(* IEC 61131-3 sources: SortJet_MasterSPS_Aufbau.fbsproj/09_Station/Stationen/Faecherwagen [301-305], 6 files *)

(* ---- I_Faecherwagenstation.itf ---- *)
(* METADATA
{
	"v3Meta": {
		"objectGuid": "03e38843-2da5-4b21-8acb-320ccd699887"
	}
}
*)
INTERFACE I_Faecherwagenstation EXTENDS __System.IQueryInterface
END_INTERFACE

(* ---- Basic_Faecherwagenstation_FB_V01_00_00.fb.st ---- *)
(* METADATA
{
	"v3Meta": {
		"objectGuid": "908407cd-758c-45db-8a2d-c326aeb0e347"
	}
}
*)
FUNCTION_BLOCK ABSTRACT Basic_Faecherwagenstation_FB_V01_00_00 EXTENDS Basic_Station_FB_V01_00_00 IMPLEMENTS I_Faecherwagenstation
VAR_INPUT

  // BOOL
  blMerkerEinschleusenQuittiert     : BOOL; // Einschleusen vom Bediener an der Station quittiert
  bpRolltorUnten                    : BOOL; // Rolltor unten (aus der Sicherheitstechnik)
  bpMMIFWBaldVoll                   : BOOL; // Faecherwagen in der Station laut MMI bald voll (Anzeige an der Station), Ruecksetzen beim Verlassen der Beladeposition

  // WORD
  wlRFID_Nummer_Schreiben           : WORD; // Neue Nummer fuer den RFID-Chip des Faecherwagens (vom MMI)

  // USINT
  usilErrorSafety                   : USINT; // Fehlercode der sicheren Feldbox (Schmersal), im Geraetebaum gemappt

END_VAR
VAR_OUTPUT

  // BOOL
  bpDone                            : BOOL;
  bpEinschleusenAbgeschlossen       : BOOL;
  bpAusschleusenAbgeschlossen       : BOOL;
  bpAuftragAktiv                    : BOOL;
  bpFehler                          : BOOL;
  bpErzwingeAusschleusen            : BOOL;
  bpErzwingeEinschleusen            : BOOL;
  bpBoxInHomePosition               : BOOL; // Mechanik der Station in Grundstellung
  bpOutBereitZumAustransport        : BOOL; // OUT STATUS: Bereit zum Austransport [Eintransport auf die Nachfolgerstation]
  bpOutBereitZumEintransport        : BOOL; // OUT STATUS: Bereit zum Eintransport [Austransport auf die Vorgaengerstation]
  bpStatusStationInBeladePosition   : BOOL; // Faecherwagen steht in der Beladeposition (zyklisch)
  bpHinweisEingriffErforderlich     : BOOL; // Bedienereingriff am Faecherwagen erforderlich (Ampel blau blinkend, Aktion Ampelsignal in Job)

  // WORD
  wpFehlerNr                        : Fehlerkonstanten_EN; // FEHLER-AUSWERTUNG: Fehlernummer[Const]

END_VAR
VAR

  // BOOL
  blRolltorAuf                      : BOOL; // Anforderung Rolltor oeffnen
  blRolltorAb                       : BOOL; // Anforderung Rolltor schliessen
  blRolltorAufDone                  : BOOL;
  blRolltorAbDone                   : BOOL;
  blRolltorAbFreigabe               : BOOL := TRUE; // Variante: Rolltor darf schliessen (z.B. nichts im Bereich des Rolltors)
  blRolltorAbBlockiert              : BOOL; // Variante: Schliessen sofort mit Fehler abbrechen (z.B. Abrollsicherung ausgeloest)
  blStationsposUndefiniert          : BOOL; // Station weder in Grundstellung noch in Beladeposition und kein Auftrag aktiv
  blStarteSicherheitskreisReset     : BOOL; // Anforderung Sicherheitsrelais der Station quittieren (MMI, Variante setzt nach Ausfuehrung zurueck)
  blAckRequested                    : BOOL; // Sichere Feldbox fordert Quittierung an, im Geraetebaum gemappt
  blResetSchmersal                  : BOOL; // Quittierimpuls an die sichere Feldbox, im Geraetebaum gemappt

  // WORD
  wlZeitHochfahren                  : WORD;
  wlZeitRunterfahren                : WORD;
  wlRFID_Nummer                     : WORD; // Zuletzt gelesene RFID-Nummer des Faecherwagens

  // TIME
  tlZeitHochfahren                  : TIME;
  tlZeitRunterfahren                : TIME;

  // STEPS
  steplRolltorAuf                   : Steps_TE;
  steplRolltorAb                    : Steps_TE;

  // TIMER
  tonlFreigabe                      : TON;
  tonlUeberwachungRolltor           : TON;
  tonlRolltorOeffnenSchliesen       : TON;
  tonlZeitRunterfahren              : TON; // Zum ermitteln wie lange das Rolltor runterfaehrt
  tonlZeitHochfahren                : TON; // Zum ermitteln wie lange das Rolltor hochfaehrt
  tplResetSchmersal                 : TP;

  // TRIGGER
  rtlSafetyError                    : R_TRIG;

  // ENUM
  eLetzterStatus                    : eLetzter_FW_Status; // Zuletzt erreichter Schritt fuer Systemcheck und MMI
  elLetzterStatusGesendet           : eLetzter_FW_Status; // Zuletzt ans MMI gemeldeter Status (STATION_UPDATE)

  // HARDWARE: ROLLTOR
  in_bRolltorGeoeffnet                     : BOOL; // TRUE = Rolltor oben, im Geraetebaum gemappt
  out_bRolltorAb                    AT %Q* : BOOL;
  out_bRolltorAuf                   AT %Q* : BOOL;

  // HARDWARE: SICHERHEITSKREIS DER STATION (im Geraetebaum gemappt)
  in_bResetSicherheitskreis         : BOOL; // Taster Sicherheitskreis quittieren an der Station
  out_bSicherheitskreisAusgeloest   : BOOL; // Leuchte Sicherheitskreis ausgeloest (Variante darf ueberschreiben)

END_VAR
VAR CONSTANT

  // TIME
  cZEIT_UEBERWACHUNG_ROLLTOR        : TIME := T#60S;

END_VAR
//-------------------------------------------------------------------------------------------------
// MASTER AUFRUFEN
//-------------------------------------------------------------------------------------------------
IF NOT __ISVALIDREF(BasisStationsParameter.stMKs) THEN
  dwpHandfunktionenReturn := DWORD#0;
  RETURN;
END_IF

SUPER^(BasisStationsParameter := BasisStationsParameter);

//-------------------------------------------------------------------------------------------------
// DEAKTIVIEREN
//-------------------------------------------------------------------------------------------------
// Werte wieder passend abloeschen, wenn der Baustein wieder aktiviert wird
IF ( ftlBausteinDeaktivierung.Q ) THEN
  bpDone                      := FALSE;
  bpEinschleusenAbgeschlossen := FALSE;
  bpAusschleusenAbgeschlossen := FALSE;
END_IF

(* Hinweis:
   - Deaktivierte Station: nichts melden, nichts bewegen
   - Die Variante prueft die Deaktivierung nach dem Aufruf selbst und setzt ihre Anforderungen zurueck
*)
IF ( BasisStationsParameter.stMKs.bDeaktivieren ) THEN

  bpDone                          := TRUE;
  bpEinschleusenAbgeschlossen     := TRUE;
  bpAusschleusenAbgeschlossen     := TRUE;
  bpStatusStationInBeladePosition := FALSE;
  bpAuftragAktiv                  := FALSE;
  bpFehler                        := FALSE;
  blStationsposUndefiniert        := FALSE;

  blRolltorAuf                    := FALSE;
  blRolltorAb                     := FALSE;
  out_bRolltorAuf                 := FALSE;
  out_bRolltorAb                  := FALSE;

  A_Visu();
  RETURN;

END_IF

//-------------------------------------------------------------------------------------------------
// TIMER
//-------------------------------------------------------------------------------------------------
tonlFreigabe( IN := BasisStationsParameter.stFreigabe.bAlles, PT := T#1S );

bpFehler := BasisStationsParameter.bFehler;

//-------------------------------------------------------------------------------------------------
// SICHERE FELDBOX / SICHERHEITSKREIS
//-------------------------------------------------------------------------------------------------
rtlSafetyError( CLK := usilErrorSafety <> 0 );
IF rtlSafetyError.Q THEN

  SpsError( eFehler_Safety_Schmersal,
            usilErrorSafety,
            BasisStationsParameter.stMKs.stStationsNummern.NummerIntern,
            AutomatikkreisBestimmen(BasisStationsParameter.stMKs.stStationsNummern.NummerSPS),
            BasisStationsParameter.awFehlerInformationen );

END_IF

tplResetSchmersal( IN := blAckRequested XOR ( NotHalt.in_bTasterNothaltQuittieren OR in_bResetSicherheitskreis ),
                   PT := T#500MS,
                   Q  => blResetSchmersal );

// Meldung "Faecherwagen bald voll" gilt nur fuer den Faecherwagen in der Beladeposition
IF NOT bpStatusStationInBeladePosition THEN
  bpMMIFWBaldVoll := FALSE;
END_IF

//-------------------------------------------------------------------------------------------------
// STATUS AN MMI MELDEN
//-------------------------------------------------------------------------------------------------
// Hinweis:
//   - Der fuer den Systemcheck gemerkte Status (eLetzterStatus) wird bei jeder Aenderung und bei
//     neuer MMI-Verbindung gemeldet; das MMI zeigt die Geraete der Station passend dazu an
IF ( eLetzterStatus <> elLetzterStatusGesendet ) OR Job.rtlMmiOk.Q THEN
  stStationUpdate.wStationsNummer       := BasisStationsParameter.stMKs.stStationsNummern.NummerSPS;
  stStationUpdate.eUpdateTyp            := StationUpdateTyp_EN.FW_STATUS;
  stStationUpdate.wAnzahlWerte          := 1;
  stStationUpdate.astWerte[1].eDatenTyp := UpdateDatenTyp_EN.TYP_WORD;
  stStationUpdate.astWerte[1].wWert     := TO_WORD( eLetzterStatus );
  MsgToMmi( auftragsnr_w := SB0_SPS_STATION_UPDATE );

  elLetzterStatusGesendet := eLetzterStatus;
END_IF
END_FUNCTION_BLOCK

(* ---- Faecherwagenstation_Einfach_FB_V01_00_00.fb.st ---- *)
(* METADATA
{
	"v3Meta": {
		"objectGuid": "602268ae-05d1-404e-8d8e-505fe92152ba"
	}
}
*)
FUNCTION_BLOCK Faecherwagenstation_Einfach_FB_V01_00_00 EXTENDS Basic_Faecherwagenstation_FB_V01_00_00
VAR_INPUT

  // BOOL
  bpFaecherwagenVorhanden          : BOOL; // Faecherwagen vorhanden, Sicherheitssensor ueber die SLC (Interface_SLC)
  in_bDruckluftOK                  : BOOL;

END_VAR
VAR

  // BOOL
  blArretierungSchliessen          : BOOL; // Anforderung Arretierung ausfahren (Faecherwagen festhalten)
  blArretierungOeffnen             : BOOL; // Anforderung Arretierung einfahren (Faecherwagen freigeben)
  blArretierungSchliessenDone      : BOOL;
  blArretierungOeffnenDone         : BOOL;
  blArretierungGeschlossen         : BOOL; // Arretierung ausgefahren (Endlage)
  blArretierungOffen               : BOOL; // Arretierung eingefahren (Endlage)
  blHandFreigabe                   : BOOL; // Handfunktionen nur im Handbetrieb zulassen
  blTasterLeuchteAnforderung       : BOOL;

  // WORD
  wlIoccMeldungsNummer             : WORD;

  // STEPS
  steplEinschleusen                : Steps_TE;
  steplAusschleusen                : Steps_TE;

  // TIMER
  tonlFWInBox                      : TON; // Faecherwagen steht stabil in der Station
  tonlErzwungenesAuschleusen       : TON;

  // TRIGGER
  rtlLogIn                         : R_TRIG;
  rtlQuittierungEinschleusen       : R_TRIG;
  rtlBetriebsartHand               : R_TRIG;
  ftlBetriebsartAutomatik          : F_TRIG;
  rtlArretierungFehler             : R_TRIG;

  // BAUSTEINE
  Arretierung                      : Arretierung_FB_V01_00_00; // Arretierung (Zentrierung/Klemmung) des ganzen Faecherwagens

  // HARDWARE EINGAENGE (Konfiguration_FW_Einfach)
  in_bAbrollsicherungOK            AT %I* : BOOL; // Abrollsicherung am Rolltor in Ordnung (Oeffner: TRUE = frei)

  // HARDWARE EINGAENGE (IO-Link, im Geraetebaum gemappt)
  in_bArretierungAusgefahren       : BOOL; // Faecherwagen arretiert
  in_bArretierungEingefahren       : BOOL; // Faecherwagen freigegeben
  in_bStartSchleusen               : BOOL; // Taster Ein-/Ausschleusen an der Station

  // HARDWARE AUSGAENGE (IO-Link, im Geraetebaum gemappt)
  out_bArretierungAusfahren        : BOOL;
  out_bArretierungEinfahren        : BOOL;
  out_bFreigabeSchleusen           : BOOL; // Leuchte im Taster Ein-/Ausschleusen

END_VAR
VAR CONSTANT

  // TIME
  ZEIT_ZWANGSAUSSCHLEUSEN          : TIME := T#3S;
  ZEIT_FW_IN_BOX                   : TIME := T#2S;

END_VAR

//-------------------------------------------------------------------------------------------------
// MASTER AUFRUFEN
//-------------------------------------------------------------------------------------------------
IF NOT __ISVALIDREF(BasisStationsParameter.stMKs) THEN
  dwpHandfunktionenReturn := DWORD#0;
  RETURN;
END_IF

SUPER^(BasisStationsParameter := BasisStationsParameter);

//-------------------------------------------------------------------------------------------------
// DEAKTIVIEREN
//-------------------------------------------------------------------------------------------------
IF ( BasisStationsParameter.stMKs.bDeaktivieren ) THEN

  blArretierungSchliessen   := FALSE;
  blArretierungOeffnen      := FALSE;
  out_bArretierungAusfahren := FALSE;
  out_bArretierungEinfahren := FALSE;
  out_bFreigabeSchleusen    := FALSE;

  HandfunktionenStatus();
  RETURN;

END_IF

//-------------------------------------------------------------------------------------------------
// AKTIONEN
//-------------------------------------------------------------------------------------------------
A_Eingaenge();
Ausschleusen();
Einschleusen();
Rolltor();

Systemcheck();

Reset();
Handfunktionen();

A_Aufrufe();
Ausgaenge();

A_Visu();
A_VisuVariante();

//-------------------------------------------------------------------------------------------------
// TASTER
//-------------------------------------------------------------------------------------------------
IF BasisStationsParameter.bEintransport[cWAND_1] THEN

  IF steplEinschleusen = STEP_105_E THEN
    blTasterLeuchteAnforderung := gbFlashbit05sec; // Einschleusen wartet auf die Quittierung
  ELSE
    blTasterLeuchteAnforderung := gbFlashbit1sec;
  END_IF

ELSIF BasisStationsParameter.bAustransport[cWAND_1] THEN
  blTasterLeuchteAnforderung := gbFlashbit1sec;

ELSIF blStationsposUndefiniert THEN
  blTasterLeuchteAnforderung := gbFlashbit02sec; // Undefinierter Zustand - sehr schnell blinken

ELSIF bpStatusStationInBeladePosition THEN
  blTasterLeuchteAnforderung := bpMMIFWBaldVoll; // Faecherwagen in Beladeposition: Dauerlicht, wenn er laut MMI bald voll ist

ELSIF bpBoxInHomePosition THEN
  blTasterLeuchteAnforderung := TRUE; // Station bereit zum Einschleusen

ELSE
  blTasterLeuchteAnforderung := gbFlashbit02sec;
END_IF

out_bFreigabeSchleusen := blTasterLeuchteAnforderung;

//-------------------------------------------------------------------------------------------------
// GESONDERTE LOGIK
//-------------------------------------------------------------------------------------------------

// Ausschleusen erzwingen: Taster lange druecken
tonlErzwungenesAuschleusen( IN := in_bStartSchleusen, PT := ZEIT_ZWANGSAUSSCHLEUSEN );
bpErzwingeAusschleusen := tonlErzwungenesAuschleusen.Q;

// Faecherwagen anmelden: Taster bei Faecherwagen in der Station und Station in Grundstellung
rtlLogIn( CLK :=     in_bStartSchleusen
                 AND bpBoxInHomePosition
                 AND tonlFWInBox.Q
                 AND NOT bpStatusStationInBeladePosition
                 AND NOT bpAuftragAktiv );

IF ( rtlLogIn.Q ) THEN
  wSps2FaecherwagenStationNr              := BasisStationsParameter.stMKs.stStationsNummern.NummerSPS;
  tMmi2SpsInfo.wSps2FaecherwagenStationNr := BasisStationsParameter.stMKs.stStationsNummern.NummerSPS;
  MsgToMmi( auftragsnr_w := SB0_SPS_RACKLOGIN );

  M_SB0_MMI_RELEASERACKLOGIN    := TRUE;
  blMerkerEinschleusenQuittiert := TRUE;
END_IF
END_FUNCTION_BLOCK

(* ---- Faecherwagenstation_Hydraulik_FB_V01_00_00.fb.st ---- *)
(* METADATA
{
	"v3Meta": {
		"objectGuid": "e6879d41-371d-40de-a0ee-fe2898e6d6d8"
	}
}
*)
FUNCTION_BLOCK Faecherwagenstation_Hydraulik_FB_V01_00_00 EXTENDS Basic_Faecherwagenstation_FB_V01_00_00
VAR_OUTPUT

  // BOOL
  bpAnforderungHydraulikEin        : BOOL; // Hydraulikaggregat einschalten (eine hydraulische Bewegung ist angefordert)
  bpUmlaufVentilPause              : BOOL; // Umlaufventil zwischen zwei direkt folgenden Bewegungen kurz zuruecknehmen

END_VAR
VAR

  // BOOL: Anforderungen
  blHubrahmenHeben                 : BOOL;
  blHubrahmenSenken                : BOOL;
  blFaecherwagenVor                : BOOL;
  blFaecherwagenZurueck            : BOOL;
  blZentrierungOeffnen             : BOOL;
  blZentrierungSchliessen          : BOOL;
  blAnschlagAuf                    : BOOL;
  blAnschlagAb                     : BOOL;
  blAnschlagVor                    : BOOL; // Option AGV: Anschlag nach vorne
  blAnschlagZurueck                : BOOL; // Option AGV: Anschlag nach hinten

  // BOOL: Bewegungen abgeschlossen
  blHubrahmenHebenDone             : BOOL;
  blHubrahmenSenkenDone            : BOOL;
  blFaecherwagenVorDone            : BOOL;
  blFaecherwagenZurueckDone        : BOOL;
  blZentrierungOeffnenDone         : BOOL;
  blZentrierungSchliessenDone      : BOOL;
  blAnschlagAufDone                : BOOL;
  blAnschlagAbDone                 : BOOL;
  blAnschlagVorDone                : BOOL;
  blAnschlagZurueckDone            : BOOL;

  // BOOL: Verschiedenes
  blFaecherwagenErkannt            : BOOL; // Beide Muting-Sensoren belegt
  blAnschlagUntenOderOhne          : BOOL; // Anschlag unten oder kein Anschlag laut MK
  blLadepositionOhneOben           : BOOL; // Beladeposition bis auf den abgesackten Hubrahmen
  blPositionskorrekturAktiv        : BOOL; // Hubrahmen wird nachgehoben
  blAnforderungHydraulik           : BOOL;
  blHandFreigabe                   : BOOL; // Handfunktionen nur im Handbetrieb zulassen
  blTasterLeuchteAnforderung       : BOOL;
  blHydraulikLaeuft                : BOOL; // Rueckmeldung der zugeordneten Hydraulikstation
  blStationBeladen                 : BOOL; // Faecherwagen eingeschleust (Status fuer AGV-Betrieb)
  blStartUp                        : BOOL := TRUE; // Sicherheitsrelais nach dem Programmstart einmal quittieren

  // BOOL: Begrenzung gleichzeitiger Auftraege je Hydraulikstation
  blHydraulikAuftragAnfrage        : BOOL; // Kette wartet auf die Freigabe eines neuen Auftrags (je Zyklus neu gesetzt)
  blHydraulikAuftragFreigabe       : BOOL; // Rueckmeldung der Hydraulikstation (M_AuftragFreigabe, letzter Zyklus)
  blHydraulikAuftragAktiv          : BOOL; // Ein-/Ausschleusen mit hydraulischen Bewegungen laeuft, belegt die Hydraulikstation
  blAuftragWartetAufHydraulik      : BOOL; // Auftrag erteilt, Hydraulikstation laesst noch keinen weiteren Auftrag zu

  // BOOL: Muting
  blMutingAusschalten              : BOOL; // Option AGV: Muting dauerhaft zuruecksetzen (kein Faecherwagen eingeschleust)
  blMutingResetAnforderung         : BOOL; // Anforderung Muting-Sensoren zuruecksetzen pruefen
  blMutingResetImpuls              : BOOL; // Reset-Impuls fuer die Muting-Sensoren ausgeben
  blMutingSensorReset              : BOOL; // Reset-Impuls aktiv

  // BYTE
  bylRFID_Nummer                   : BYTE;

  // WORD
  wlIoccMeldungsNummer             : WORD;
  wlStationStatusWord              : WORD; // Option AGV: zuletzt ans MMI gemeldeter Status der Station

  // REFERENZ
  refHydraulikstation              : REFERENCE TO Hydraulik_FB_V01_00_00; // laut MK stStationsAufbau.wHydraulikstation

  // STEPS
  steplEinschleusen                : Steps_TE;
  steplAusschleusen                : Steps_TE;
  steplHubrahmenHeben              : Steps_TE;
  steplHubrahmenSenken             : Steps_TE;
  steplFaecherwagenVor             : Steps_TE;
  steplFaecherwagenZurueck         : Steps_TE;
  steplZentrierungOeffnen          : Steps_TE;
  steplZentrierungSchliessen       : Steps_TE;
  steplSicherheitskreisReset       : Steps_TE;

  // TIMER
  tonlHubrahmenUeberfahren         : TON; // Sensor ueberfahren, Endlage sicher erreicht
  tonlVerfahrenUeberfahren         : TON;
  tonlZentrierungUeberfahren       : TON;
  tonlTimeoutHubrahmen             : TON;
  tonlTimeoutVerfahren             : TON;
  tonlTimeoutZentrierung           : TON;
  tonlTimeoutHydraulik             : TON; // Warten auf das Hydraulikaggregat
  tonlTimeoutReadRFID              : TON;
  tonlFWInBox                      : TON;
  tonlErzwungenesAuschleusen       : TON;
  tonlMutingSensorFehler           : TON;
  tonlPositionskorrektur           : TON;
  tonlUmlaufventilPause            : TON; // Dauer der Pause des Umlaufventils
  tonlMutingSensorenBelegt         : TON; // Beide Muting-Sensoren stabil belegt
  tonlTimeoutAGV                   : TON; // Option AGV: Warten auf den Faecherwagen
  tonlRFIDGelesen                  : TON; // Option AGV: RFID-Chip stabil gelesen
  tonlStartUp                      : TON;
  tonlResetImpuls                  : TON; // Impulsdauer Reset Sicherheitsrelais
  tonlResetWarten                  : TON; // Wartezeiten der Kette Sicherheitskreis-Reset
  toflAnforderungHydraulikEin      : TOF;
  toflMutingSensorReset            : TOF; // Impulsdauer Reset Muting-Sensoren

  // TRIGGER
  rtlLogIn                         : R_TRIG;
  rtlQuittierungEinschleusen       : R_TRIG;
  rtlBetriebsartHand               : R_TRIG;
  ftlBetriebsartAutomatik          : F_TRIG;
  rtlPositionskorrektur            : R_TRIG;
  rtlAnschlagFehler                : R_TRIG;
  rtlAnschlagHorizontalFehler      : R_TRIG;
  rtlMutingSensorReset             : R_TRIG;
  ftlRFIDNichtMehrGelesen          : F_TRIG;

  // BAUSTEINE
  Anschlag                         : ZylinderPneumatik_FB_V01_00_00; // Option stStationsAufbau.bAnschlag, ausgefahren = oben
  AnschlagHorizontal               : ZylinderPneumatik_FB_V01_00_00; // Option bAnschlag und bAGV, ausgefahren = vorne

  // HARDWARE EINGAENGE
  in_bHubrahmenOben                AT %I* : BOOL;
  in_bHubrahmenUnten               AT %I* : BOOL;
  in_bFaecherwagenVorne            AT %I* : BOOL;
  in_bFaecherwagenHinten           AT %I* : BOOL;
  in_bZentrierungOffen             AT %I* : BOOL;
  in_bZentrierungGeschlossen       AT %I* : BOOL;
  in_bAnschlagOben                 AT %I* : BOOL;
  in_bAnschlagUnten                AT %I* : BOOL;
  in_bAnschlagVorne                AT %I* : BOOL; // Option AGV
  in_bAnschlagHinten               AT %I* : BOOL; // Option AGV
  in_bFWInAusrichtPosition         AT %I* : BOOL; // Faecherwagen steht vor der Station in Ausrichtposition
  in_bMutingSensorLinks            AT %I* : BOOL;
  in_bMutingSensorRechts           AT %I* : BOOL;
  in_bStartSchleusen               AT %I* : BOOL; // Taster Ein-/Ausschleusen an der Station
  in_bSicherheitsrelaisOK          AT %I* : BOOL;
  in_bAbrollsicherungOK            AT %I* : BOOL; // Abrollsicherung des Rolltors nicht ausgeloest
  in_bRFID_DataValid               AT %I* : BOOL;
  in_bRFID_NR1                     AT %I* : BOOL;
  in_bRFID_NR2                     AT %I* : BOOL;
  in_bRFID_NR3                     AT %I* : BOOL;
  in_bRFID_NR4                     AT %I* : BOOL;
  in_bRFID_NR5                     AT %I* : BOOL;
  in_bRFID_NR6                     AT %I* : BOOL;
  in_bRFID_NR7                     AT %I* : BOOL;
  in_bRFID_NR8                     AT %I* : BOOL;

  // HARDWARE AUSGAENGE
  out_bHubrahmenHeben              AT %Q* : BOOL;
  out_bHubrahmenSenken             AT %Q* : BOOL;
  out_bFaecherwagenVor             AT %Q* : BOOL;
  out_bFaecherwagenZurueck         AT %Q* : BOOL;
  out_bZentrierungOeffnen          AT %Q* : BOOL;
  out_bZentrierungSchliessen       AT %Q* : BOOL;
  out_bAnschlagAuf                 AT %Q* : BOOL;
  out_bAnschlagAb                  AT %Q* : BOOL;
  out_bAnschlagVor                 AT %Q* : BOOL; // Option AGV
  out_bAnschlagZurueck             AT %Q* : BOOL; // Option AGV
  out_bFreigabeSchleusen           AT %Q* : BOOL; // Leuchte im Taster Ein-/Ausschleusen
  out_bMutingSensorReset           AT %Q* : BOOL; // Muting-Sensoren zuruecksetzen
  out_bResetSicherheitsrelais      AT %Q* : BOOL; // Sicherheitsrelais der Station quittieren

END_VAR
VAR CONSTANT

  // TIME
  ZEIT_TIMEOUT_SENSOR              : TIME := T#30S;
  ZEIT_TIMEOUT_HYDRAULIK           : TIME := T#30S;
  ZEIT_SENSOR_UEBERFAHREN          : TIME := T#3S;
  ZEIT_POSITIONSKORREKTUR          : TIME := T#5S;
  ZEIT_TIMEOUT_RFID                : TIME := T#5S;
  ZEIT_ZWANGSAUSSCHLEUSEN          : TIME := T#3S;
  ZEIT_FW_IN_BOX                   : TIME := T#1S;
  ZEIT_UMLAUFVENTIL_PAUSE          : TIME := T#1S;
  ZEIT_MUTING_SENSOR_RESET         : TIME := T#500MS;
  ZEIT_STARTUP_SICHERHEITSRELAIS   : TIME := T#5S;

END_VAR
//-------------------------------------------------------------------------------------------------
// MASTER AUFRUFEN
//-------------------------------------------------------------------------------------------------
IF NOT __ISVALIDREF(BasisStationsParameter.stMKs) THEN
  dwpHandfunktionenReturn := DWORD#0;
  RETURN;
END_IF

SUPER^(BasisStationsParameter := BasisStationsParameter);

//-------------------------------------------------------------------------------------------------
// DEAKTIVIEREN
//-------------------------------------------------------------------------------------------------
IF ( BasisStationsParameter.stMKs.bDeaktivieren ) THEN

  blHubrahmenHeben           := FALSE;
  blHubrahmenSenken          := FALSE;
  blFaecherwagenVor          := FALSE;
  blFaecherwagenZurueck      := FALSE;
  blZentrierungOeffnen       := FALSE;
  blZentrierungSchliessen    := FALSE;
  blAnschlagAuf              := FALSE;
  blAnschlagAb               := FALSE;
  blAnschlagVor              := FALSE;
  blAnschlagZurueck          := FALSE;
  blPositionskorrekturAktiv  := FALSE;
  blMutingResetImpuls        := FALSE;
  steplSicherheitskreisReset := STEP_0_E;

  out_bHubrahmenHeben        := FALSE;
  out_bHubrahmenSenken       := FALSE;
  out_bFaecherwagenVor       := FALSE;
  out_bFaecherwagenZurueck   := FALSE;
  out_bZentrierungOeffnen    := FALSE;
  out_bZentrierungSchliessen := FALSE;
  out_bAnschlagAuf           := FALSE;
  out_bAnschlagAb             := FALSE;
  out_bAnschlagVor            := FALSE;
  out_bAnschlagZurueck        := FALSE;
  out_bFreigabeSchleusen      := FALSE;
  out_bMutingSensorReset      := FALSE;
  out_bResetSicherheitsrelais := FALSE;
  bpAnforderungHydraulikEin   := FALSE;
  bpUmlaufVentilPause         := FALSE;

  HandfunktionenStatus();
  RETURN;

END_IF

//-------------------------------------------------------------------------------------------------
// AKTIONEN
//-------------------------------------------------------------------------------------------------
A_Eingaenge();
Ausschleusen();
Einschleusen();
Positionskorrektur();

Hubrahmen();
Verfahren();
Zentrierung();
Rolltor();

Systemcheck();
Status_Meldung();

Reset();
Handfunktionen();

MutingSensorReset();
Sicherheitskreis_Reset();

A_Aufrufe();
Ausgaenge();

A_Visu();
A_VisuVariante();

//-------------------------------------------------------------------------------------------------
// TASTER
//-------------------------------------------------------------------------------------------------
IF blAuftragWartetAufHydraulik THEN
  blTasterLeuchteAnforderung := gbFlashbit02sec; // Auftrag erteilt, wartet auf die Hydraulikstation - sehr schnell blinken

ELSIF BasisStationsParameter.bEintransport[cWAND_1] THEN

  IF steplEinschleusen = STEP_100_E THEN
    blTasterLeuchteAnforderung := gbFlashbit05sec; // Einschleusen wartet auf die Quittierung
  ELSE
    blTasterLeuchteAnforderung := gbFlashbit1sec;
  END_IF

ELSIF BasisStationsParameter.bAustransport[cWAND_1] THEN
  blTasterLeuchteAnforderung := gbFlashbit1sec;

ELSIF blStationsposUndefiniert THEN
  blTasterLeuchteAnforderung := gbFlashbit02sec; // Undefinierter Zustand - sehr schnell blinken

ELSIF bpStatusStationInBeladePosition THEN
  blTasterLeuchteAnforderung := bpMMIFWBaldVoll; // Faecherwagen in Beladeposition: Dauerlicht, wenn er laut MMI bald voll ist

ELSIF bpBoxInHomePosition AND in_bFWInAusrichtPosition THEN
  blTasterLeuchteAnforderung := TRUE; // Faecherwagen steht bereit zum Einschleusen

ELSE
  blTasterLeuchteAnforderung := FALSE;
END_IF

out_bFreigabeSchleusen := blTasterLeuchteAnforderung;

//-------------------------------------------------------------------------------------------------
// GESONDERTE LOGIK
//-------------------------------------------------------------------------------------------------

// Ausschleusen erzwingen: Taster lange druecken
tonlErzwungenesAuschleusen( IN := in_bStartSchleusen, PT := ZEIT_ZWANGSAUSSCHLEUSEN );
bpErzwingeAusschleusen := tonlErzwungenesAuschleusen.Q;

// Faecherwagen anmelden: Taster bei Faecherwagen in Ausrichtposition und Station in Grundstellung
rtlLogIn( CLK :=     in_bStartSchleusen
                 AND bpBoxInHomePosition
                 AND tonlFWInBox.Q
                 AND NOT bpStatusStationInBeladePosition
                 AND NOT bpAuftragAktiv );

IF ( rtlLogIn.Q ) THEN
  wSps2FaecherwagenStationNr              := BasisStationsParameter.stMKs.stStationsNummern.NummerSPS;
  tMmi2SpsInfo.wSps2FaecherwagenStationNr := BasisStationsParameter.stMKs.stStationsNummern.NummerSPS;
  MsgToMmi( auftragsnr_w := SB0_SPS_RACKLOGIN );

  M_SB0_MMI_RELEASERACKLOGIN    := TRUE;
  blMerkerEinschleusenQuittiert := TRUE;
END_IF

// Hydraulikaggregat einschalten, solange eine hydraulische Bewegung angefordert und nicht fertig ist
blAnforderungHydraulik :=     BasisStationsParameter.stFreigabe.bAlles
                          AND (    ( blHubrahmenHeben        AND NOT blHubrahmenHebenDone )
                                OR ( blHubrahmenSenken       AND NOT blHubrahmenSenkenDone )
                                OR ( blFaecherwagenVor       AND NOT blFaecherwagenVorDone )
                                OR ( blFaecherwagenZurueck   AND NOT blFaecherwagenZurueckDone )
                                OR ( blZentrierungOeffnen    AND NOT blZentrierungOeffnenDone )
                                OR ( blZentrierungSchliessen AND NOT blZentrierungSchliessenDone ) );

toflAnforderungHydraulikEin( IN := blAnforderungHydraulik, PT := T#2S );
bpAnforderungHydraulikEin := toflAnforderungHydraulikEin.Q;

// Anforderung an die zugeordnete Hydraulikstation melden (Aufruf der Hydraulikstation nach den Faecherwagenstationen)
IF __ISVALIDREF(refHydraulikstation) THEN
  refHydraulikstation.M_Anfordern( bpHydraulikEin      := bpAnforderungHydraulikEin,
                                   bpUmlaufventilPause := bpUmlaufVentilPause );
  blHydraulikLaeuft := refHydraulikstation.bpHydraulikLaeuft;
ELSE
  // Keine Hydraulikstation zugeordnet: hydraulische Bewegungen laufen in die Zeitueberwachung
  blHydraulikLaeuft := FALSE;
END_IF

// Begrenzung gleichzeitiger Auftraege je Hydraulikstation (MK wMaximaleAnzahlAktiverAuftraege):
// Auftrag belegt die Hydraulikstation, bis Ein-/Austransport beendet oder abgebrochen ist
IF     NOT BasisStationsParameter.bEintransport[cWAND_1]
   AND NOT BasisStationsParameter.bAustransport[cWAND_1]
THEN
  blHydraulikAuftragAktiv := FALSE;
END_IF

IF __ISVALIDREF(refHydraulikstation) THEN
  blHydraulikAuftragFreigabe := refHydraulikstation.M_AuftragFreigabe( bpAuftragAktiv   := blHydraulikAuftragAktiv OR blPositionskorrekturAktiv,
                                                                       bpAuftragStarten := blHydraulikAuftragAnfrage );
ELSE
  // Keine Hydraulikstation zugeordnet: keine Begrenzung
  blHydraulikAuftragFreigabe := TRUE;
END_IF

blAuftragWartetAufHydraulik := blHydraulikAuftragAnfrage AND NOT blHydraulikAuftragFreigabe;
blHydraulikAuftragAnfrage   := FALSE;

// Sicherheitsrelais der Station nach dem Programmstart einmal quittieren, sobald Not-Halt in Ordnung ist
tonlStartUp( IN := blStartUp AND NotHalt.bpNotHaltOK, PT := ZEIT_STARTUP_SICHERHEITSRELAIS );

IF ( tonlStartUp.Q ) THEN
  blStartUp                     := FALSE;
  blStarteSicherheitskreisReset := TRUE;
END_IF
END_FUNCTION_BLOCK

(* ---- Faecherwagenstation_Lineareinheit_FB_V01_00_00.fb.st ---- *)
(* METADATA
{
	"v3Meta": {
		"objectGuid": "3779c208-854f-4c13-8b26-aa1147fe8cdb"
	}
}
*)
FUNCTION_BLOCK Faecherwagenstation_Lineareinheit_FB_V01_00_00 EXTENDS Basic_Faecherwagenstation_FB_V01_00_00
VAR_INPUT

  // BOOL
  bpLichtschranke_OK                      : BOOL;// Eingang aus der Sicherheitsteechnik das die Lichtschrnake quittiert ist
  bpUntergestellErkannt                   : BOOL;//safety eingang der Anzeigt, ob ein Unterwagen erkannt wurde
  in_bDruckluftOK                         : BOOL;
  bpLichtschrankeWartetAufQuittierungAmOP : BOOL;

END_VAR
VAR

  //Startet eine Bewegung
  blLineareinheitVor               : BOOL;
  blLineareinheitZurueck           : BOOL;
  blLineareinheitShuttle           : BOOL;
  blEntriegelungOeffnen            : BOOL;
  blEntriegelungSchliessen         : BOOL;
  blGegenhalterOeffnen             : BOOL;
  blGegenhalterSchliessen          : BOOL;
  blGreiferOeffnen                 : BOOL;
  blGreiferSchliessen              : BOOL;
  blTagPresent                     : BOOL;

  //Bewegungen Abgeschlossen
  blLineareinheitVorDone           : BOOL;
  blLineareinheitZurueckDone       : BOOL;
  blLineareinheitShuttleDone       : BOOL;
  blEntriegelungOeffnenDone        : BOOL;
  blEntriegelungSchliessenDone     : BOOL;
  blGegenhalterOeffnenDone         : BOOL;
  blGegenhalterSchliessenDone      : BOOL;
  blGreiferOeffnenDone             : BOOL;
  blGreiferSchliessenDone          : BOOL;
  blLuftAbschaltungS1              : BOOL;
  blLuftAbschaltungS2              : BOOL;
  blVentilReset                    : BOOL;
  blLinVorBeiRolltorFahrt          : BOOL; // Einschleusen: Lineareinheit darf vorfahren, waehrend das Rolltor hochfaehrt
  blRolltorAbBeiLinZurueck         : BOOL; // Ausschleusen: Rolltor darf schliessen, waehrend die Lineareinheit zurueckfaehrt
  blOberwagenBewegenGesperrt       : BOOL; // Rolltor nicht oben + Greifer haelt Oberwagen + Lineareinheit nicht hinten/SH -> Lineareinheit darf nicht fahren
  blHandFreigabe                   : BOOL; // Handfunktionen nur im Handbetrieb zulassen

  // jeweils Zusammenfassung der beiden Eingänge
  blLinearEinheitVorne             : BOOL;
  blLinearEinheitHinten            : BOOL;
  blLinearEinheitSH                : BOOL;
  blGreiferOffen                   : BOOL;
  blGreiferZu                      : BOOL;

  //Verschiedenes
  blTasterLeuchteAnforderung       : BOOL;
  blRFID_Auslesen                  : BOOL;
  blRFID_Schreiben                 : BOOL;
  blRFID_Sensor_ModusBit_0         : BOOL;
  blRFID_Sensor_ModusBit_1         : BOOL;
  blRFID_Sensor_ModusBit_2         : BOOL;
  blRFID_Sensor_ModusBit_3         : BOOL;
  blRFID_Sensor_ModusBit_4         : BOOL;
  blRFID_Sensor_ModusBit_5         : BOOL;
  blRFID_Sensor_ModusBit_6         : BOOL;
  blRFID_Sensor_ModusBit_7         : BOOL;
  blRFID_Sensor_Write_Done         : BOOL;

  blErr1, blErr2, blErr3, blErr4, blErr5 : BOOL;

  // WORD
  wlIoccMeldungsNummer                                   : WORD;
  wlioccFWStationGegenhalterUnterwagenNichtFixiert       : WORD;
  wlioccFWStationGegenhalterUnterwagenNichtFrei          : WORD;
  wlioccFWStationRolltorNichtOben                        : WORD;
  wlioccFWStationRolltorNichtUnten                       : WORD;
  wlioccFWStationGreiferNichtGeoeffnet                   : WORD;
  wlioccFWStationGreiferNichtGeschlossen                 : WORD;
  wlioccFWStationLineareinheitNichtVorne                 : WORD;
  wlioccFWStationLineareinheitNichtHinten                : WORD;
  wlioccFWStationEntriegelungNichtGeoeffnet              : WORD;
  wlioccFWStationEntriegelungNichtGeschlossen            : WORD;
  wlioccFWStationAusrichtPositionNichtOK                 : WORD;
  wlioccStationsposUndefiniert                           : WORD;
  wlioccFWagenStationSIKreisausgeloest                   : WORD;
  wlioccFWagenStationHomeposLineareinheitNichtHinten     : WORD;
  wlioccFWagenStationHomeposGreiferNichtGeoeffnet        : WORD;
  wlioccFWagenStationHomeposRolltorNichtUnten            : WORD;
  wlioccFWagenStationHomeposEntriegelungNichtGeschlossen : WORD;
  wlioccFWagenStationHomeposGegenhalterNichtGeoeffnet    : WORD;
  wlioccFWagenStationKlemmungNichtEingefahren            : WORD;
  wlRFID_NummerMerker                                    : WORD;
  wlIndexByte                                            : WORD;
  wlIndexZiffer                                          : WORD;
  wlMaxRFIDNummer                                        : WORD;
  wlIndex_STRING                                         : WORD;
  wlioccRolltorBlockiertdurchFWNichtinPos                : WORD;

  // STEPS
  steplEinschleusen           : Steps_TE;
  steplAusschleusen           : Steps_TE;
  steplLineareinheitVor       : Steps_TE;
  steplLineareinheitZur       : Steps_TE;
  steplLineareinheitShuttle   : Steps_TE;
  steplEntriegelungOeffnen    : Steps_TE;
  steplEntriegelungSchliessen : Steps_TE;
  steplGegenhalterOeffnen     : Steps_TE;
  steplGegenhalterSchliessen  : Steps_TE;
  steplGreiferOeffnen         : Steps_TE;
  steplGreiferSchliessen      : Steps_TE;
  steplresetSIRelais          : Steps_TE;
  steplRFID_Auslesen          : Steps_TE;
  steplRFID_Schreiben         : Steps_TE;

  // TIMER
  tonlLineareinheitVorZurueck        : TON;
  tonlLineareinheitShuttle           : TON;
  tonlEntriegelungAufZu              : TON;
  tonlGegenhalterAufZu               : TON;
  tonlGreiferAufZu                   : TON;
  tonlErzwungenesAuschleusen         : TON;
  tonlFreigabeZumAusschleusen        : TON;
  tonlWagenInShuttleTransferposition : TON;
  tonlTimeoutSensorVorne             : TON;
  tonlTimeoutSensorHinten            : TON;
  tonlTimeoutSensorShutle            : TON;
  tonlTimeoutReadRFID                : TON;
  tonlTimeoutGreiferAufZu            : TON;
  tonlTimeoutGegenhalterAufZu        : TON;
  tonlTimeoutEntriegelungAufZu       : TON;
  tonlFWInBox                        : TON;
  tonlSetzeSIRealisReset             : TON;
  tonlWarteSchritt                   : TON;
  tonUntergestellErkannt             : TON;
  tofTagPresent                      : TOF;

  // TRIGGER
  rtlLogIn                           : R_TRIG;
  rtlBetriebsartHand                 : R_TRIG;
  ftlBetriebsartAutomatik            : F_TRIG;
  rtlQuittierungEinschleusen         : R_TRIG;
  rtlRFID_Schreiben                  : R_TRIG;

END_VAR

VAR

  // IO-Link-Master
  in_bLinearEinheit1Vorne         : BOOL;
  in_bLinearEinheit1Hinten        : BOOL;
  in_bLinearEinheit2Vorne         : BOOL;
  in_bLinearEinheit2Hinten        : BOOL;
  in_bFaecherwagenNichtInPos      : BOOL;
  in_bEntriegelungOffen           : BOOL;
  in_bEntriegelungGeschlossen     : BOOL;
  in_bGegenhalterOffen            : BOOL;
  in_bGegenhalterZu               : BOOL;
  in_bGreifer1Offen               : BOOL;
  in_bGreifer1Zu                  : BOOL;
  in_bKlemmZylinderEingefahren    : BOOL; //zur Fixierung des Oberrahmens beim Ein und Ausschleusen. Eingefahren = Grundstellung

  //  IO-Link-Slave
  in_bGreifer2Offen                  : BOOL;
  in_bGreifer2Zu                     : BOOL;
  out_bGreiferEinfahren              : BOOL;
  out_bGreiferAusfahren              : BOOL;
  out_bEntriegelungEinfahren         : BOOL;
  out_bEntriegelungAusfahren         : BOOL;
  in_bStartSchleusen                 : BOOL;
  out_bFreigabeSchleusen             : BOOL;
  in_bLineareinheit1Umgreifposition  : BOOL;
  in_bLineareinheit2Umgreifposition  : BOOL;
  out_bGegenhalterEinfahren          : BOOL;
  out_bGegenhalterAusfahren          : BOOL;
  out_bLinearEinheitVor              : BOOL;
  out_bLinearEinheitZurueck          : BOOL;

  blRFID_NR1                     : BOOL;
  blRFID_NR2                     : BOOL;
  blRFID_NR3                     : BOOL;
  blRFID_NR4                     : BOOL;
  blRFID_NR5                     : BOOL;
  blRFID_NR6                     : BOOL;
  blRFID_NR7                     : BOOL;
  blRFID_NR8                     : BOOL;
  blRFID_DataValid               : BOOL;
  blRFID_DataWasValid            : BOOL;

  //RFID Ansteuerung
  // Out
  out_bRFID_Sensor_Start_RW      : BOOL;
  out_bDeactivateAntenna         : BOOL;
  blCMD_END                      : BOOL;

  //tmp
  ablRFID                        : ARRAY[1..32,0..7] OF BOOL;
  ablRFID_out                                : ARRAY[1..32,0..7] OF BOOL;

  abylBytesRFID                  : ARRAY [1..32] OF BYTE; //16=R,17=a,18=c,19=k,20= ,21=0,22=0,23=9
  abylBytesRFID_out              : ARRAY [1..32] OF BYTE; //16=R,17=a,18=c,19=k,20= ,21=0,22=0,23=
  bytest                         : BYTE;

  slRFID_Nummer                  : STRING;
  slMaxRFID_Nummer               : STRING;
  slRFID_Validierung             : STRING;

END_VAR

VAR CONSTANT

  // TIME
  TIMEOUT_SENSOR           : TIME := T#2M;
  ZEIT_ZWANGSAUSSCHLEUSEN  : TIME := t#3s;
  ZEIT_MUTING_SENSOR_RESET : TIME := T#500MS;
  //String
  VERGLEICH_RFID_VALID     : STRING := 'Rack ';
  //WORD
  ERSTES_ZEICHEN           : WORD := 16;
  ERSTE_ZIFFER_RFID        : WORD := 21 ;
  ANZAHL_ZIFFERN_RFID      : WORD := 3 ;
  cByte0                   : BYTE := 0;

END_VAR

//-------------------------------------------------------------------------------------------------
// MASTER AUFRUFEN
//-------------------------------------------------------------------------------------------------
IF NOT __ISVALIDREF(BasisStationsParameter.stMKs) THEN
  dwpHandfunktionenReturn := DWORD#0;
  RETURN;
END_IF

SUPER^(BasisStationsParameter := BasisStationsParameter);

//-------------------------------------------------------------------------------------------------
// DEAKTIVIEREN
//-------------------------------------------------------------------------------------------------
IF ( BasisStationsParameter.stMKs.bDeaktivieren ) THEN

  (* Hinweis:
     - Ausgaenge zuruecksetzen
  *)
  blLineareinheitVor          := FALSE;
  blLineareinheitZurueck      := FALSE;
  blLineareinheitShuttle      := FALSE;
  blEntriegelungOeffnen       := FALSE;
  blEntriegelungSchliessen    := FALSE;
  blGegenhalterOeffnen        := FALSE;
  blGegenhalterSchliessen     := FALSE;
  blGreiferOeffnen            := FALSE;
  blGreiferSchliessen         := FALSE;

  HandfunktionenStatus();
  RETURN;

END_IF

//-------------------------------------------------------------------------------------------------
// AKTIONEN
//-------------------------------------------------------------------------------------------------
A_Eingaenge();
Entriegelung();
Ausschleusen();
Einschleusen();
Linereinheit();

// Rolltor nur schliessen, wenn die Lineareinheit nicht im Bereich des Rolltors steht
// (Ausschleusen: schon waehrend die Lineareinheit mit offenem Greifer zurueckfaehrt)
blRolltorAbFreigabe := blLinearEinheitHinten OR blLinearEinheitSH OR blRolltorAbBeiLinZurueck;
Rolltor();

Gegenhalter();
Greifer();
RFID_Auslesen();
RFID_Schreiben();

Systemcheck();

Reset();
Handfunktionen();

Ausgaenge();

A_Visu();
A_VisuVariante();

//-------------------------------------------------------------------------------------------------
// TASTER
//-------------------------------------------------------------------------------------------------

// Hiwneis:
//    - Auftrag aktiv
IF BasisStationsParameter.bEintransport[1] THEN

  IF steplEinschleusen = STEP_105_E THEN
    blTasterLeuchteAnforderung := gbFlashbit05sec; // Eintransport wartet auf Quittierung oder Lichtschranke
  ELSE
    blTasterLeuchteAnforderung := gbFlashbit1sec;
  END_IF

ELSIF BasisStationsParameter.bAustransport[1] THEN
  IF steplAusschleusen = STEP_10_E THEN
    blTasterLeuchteAnforderung := gbFlashbit05sec;
  ELSIF steplAusschleusen = STEP_143_E THEN
    blTasterLeuchteAnforderung := gbFlashbit02sec;
  ELSE
    blTasterLeuchteAnforderung := gbFlashbit1sec;
  END_IF
ELSE
  IF blStationsposUndefiniert THEN
    blTasterLeuchteAnforderung := gbFlashbit02sec; // Undefinierter Zustand - sehr schnell blinken
  ELSIF bpStatusStationInBeladePosition THEN
    blTasterLeuchteAnforderung := bpMMIFWBaldVoll; // Fächerwagen in Box: Dauerlicht, wenn er laut MMI bald voll ist, sonst aus
  ELSIF bpBoxInHomePosition THEN
    blTasterLeuchteAnforderung := TRUE; // Fächerwagenbox ist leer
  ELSE
    blTasterLeuchteAnforderung := gbFlashbit02sec; // Undefinierter Zustand - sehr schnell blinken
  END_IF
END_IF

out_bFreigabeSchleusen := blTasterLeuchteAnforderung;

//-------------------------------------------------------------------------------------------------
// GESONDERTE LOGIK
//-------------------------------------------------------------------------------------------------

(* Hinweis:
   - Ausschleusen erzwingen
*)
tonlErzwungenesAuschleusen( IN := in_bStartSchleusen, PT := ZEIT_ZWANGSAUSSCHLEUSEN );
tonlLineareinheitShuttle(IN:=blLinearEinheitSH, PT := T#2S);
bpErzwingeAusschleusen := tonlErzwungenesAuschleusen.Q;

(* Hinweis:
   - FW einschleusen
*)
tonlFWInBox(IN := blTagPresent, PT := T#2S);
tofTagPresent(IN := blTagPresent, PT := T#2S);

rtlLogIn( CLK := in_bStartSchleusen
          AND bpBoxInHomePosition
          AND bpUntergestellErkannt
          AND tonlFWInBox.Q
          AND NOT bpStatusStationInBeladePosition
          AND NOT bpAuftragAktiv );

IF ( rtlLogIn.Q ) THEN
  wSps2FaecherwagenStationNr              := BasisStationsParameter.stMKs.stStationsNummern.NummerSPS;
  tMmi2SpsInfo.wSps2FaecherwagenStationNr := BasisStationsParameter.stMKs.stStationsNummern.NummerSPS;
  MsgToMmi( auftragsnr_w := SB0_SPS_RACKLOGIN );

  M_SB0_MMI_RELEASERACKLOGIN    := TRUE;
  blMerkerEinschleusenQuittiert := TRUE;
END_IF

//-------------------------------------------------------------------------------------------------
// RFID Chip beschreiben
//-------------------------------------------------------------------------------------------------
rtlRFID_Schreiben(CLK :=wlRFID_Nummer_Schreiben > 0);
IF rtlRFID_Schreiben.Q THEN
  blRFID_Schreiben    := TRUE;
  blRFID_Auslesen     := FALSE;
END_IF

//-------------------------------------------------------------------------------------------------
// Kollision mit Rolltor verhindern
//-------------------------------------------------------------------------------------------------
// Ventil für die Lineareinheiten auf Home Pos schlaten falls das Ventiel Lineareinheit in Richtung geschlossenes Rolltor fährt
// - Wenn kein Unterwagen vorhanden ist und das Rolltor geschlossen ist sollte auch kein Oberwagen in der Anlage sein

tonUntergestellErkannt (IN:= NOT bpUntergestellErkannt, PT:= T#2S);

// Oberwagen nie bewegen (reinziehen / rausschieben), solange das Rolltor nicht oben ist und die Lineareinheit ihn haelt:
//   - Greifer nicht offen und Lineareinheit nicht in Endlage hinten / SH -> Lineareinheit steht am Oberwagen
//   - z.B. Abbruch Einschleusen (Rolltor-Timeout) nachdem die Lineareinheit am FW gegriffen hat
//   - Hat Vorrang vor dem Zwangs-Zurueck unten, Ausgaenge bleiben aus bis Rolltor oben oder Greifer offen
//   - Die mechanische Oberwagensperre schaltet gegenlaeufig zum Greifer und wird nicht eigens angesteuert
blOberwagenBewegenGesperrt :=     BasisStationsParameter.stMKs.stStationsAufbau.bRolltor
                              AND NOT in_bRolltorGeoeffnet
                              AND NOT blGreiferOffen
                              AND NOT blLinearEinheitHinten
                              AND NOT blLinearEinheitSH;

IF blOberwagenBewegenGesperrt THEN
  out_bLinearEinheitZurueck := FALSE;
  out_bLinearEinheitVor     := FALSE;
  blVentilReset             := FALSE;

ELSIF (    tonUntergestellErkannt.Q
        OR ( NOT in_bRolltorGeoeffnet AND NOT blLinVorBeiRolltorFahrt ) ) THEN // Einschleusen: Vorfahren waehrend Rolltor hochfaehrt erlaubt

  blVentilReset := TRUE;

  IF blVentilReset THEN
    out_bLinearEinheitZurueck := TRUE;
    out_bLinearEinheitVor     := FALSE;

  ELSE
    out_bLinearEinheitZurueck := FALSE;
    out_bLinearEinheitVor     := FALSE;

  END_IF
ELSE
  blVentilReset := FALSE;
END_IF
END_FUNCTION_BLOCK

(* ---- Hydraulik_FB_V01_00_00.fb.st ---- *)
(* METADATA
{
	"v3Meta": {
		"objectGuid": "c072031a-76c2-44a8-94fd-df0eea8cf4c6"
	}
}
*)
FUNCTION_BLOCK Hydraulik_FB_V01_00_00
VAR_INPUT

  // WORD
  wpHydraulikstationNr             : WORD; // Nummer der Hydraulikstation (Index in apgMKHydraulikstation)

END_VAR
VAR_OUTPUT

  // BOOL
  bpHydraulikLaeuft                : BOOL; // Aggregat laeuft, Umlaufventil geschlossen: hydraulische Bewegungen moeglich

END_VAR
VAR

  // BOOL
  blErsterZyklus                   : BOOL := TRUE;
  blAnforderungHydraulik           : BOOL; // Gesammelte Anforderungen der Faecherwagenstationen (laufender Zyklus)
  blAnforderungUmlaufventilPause   : BOOL; // Gesammelte Pausen-Anforderungen der Faecherwagenstationen (laufender Zyklus)
  blHydraulikStarten               : BOOL;
  blUmlaufventilPause              : BOOL;

  // WORD
  wlAktiveAuftraege                : WORD; // Aktive Auftraege der zugeordneten Stationen (letzter Zyklus)
  wlAktiveAuftraegeZyklus          : WORD; // Aktive Auftraege (laufender Zyklus, ueber M_AuftragFreigabe)
  wlNeueAuftraegeZyklus            : WORD; // Im laufenden Zyklus neu freigegebene Auftraege

  // REFERENZ
  refMK                            : REFERENCE TO Parameter_Hydraulikstation;

  // TIMER
  tonlUmlaufventilEin              : TON; // Umlaufventil erst nach dem Hochlaufen des Motors schalten

  // HARDWARE EINGAENGE
  in_bMotorschuetz_Hydraulikkreislauf_OK  AT %I* : BOOL;

  // HARDWARE AUSGAENGE
  out_bHydraulikkreislauf_MotorEin        AT %Q* : BOOL;
  out_bHydraulikkreislauf_UmlaufventilAuf AT %Q* : BOOL;

END_VAR
VAR CONSTANT

  // WORD
  cUMRECHNUNG_MILLISEKUNDEN_SEKUNDEN : WORD := WORD#1000;

END_VAR

//-------------------------------------------------------------------------------------------------
// INITIALISIERUNG
//-------------------------------------------------------------------------------------------------
IF ( blErsterZyklus ) THEN
  blErsterZyklus := FALSE;

  IF     ( wpHydraulikstationNr >= cERSTE_HYDRAULIKSTATIONS_NR )
     AND ( wpHydraulikstationNr <= cLETZTE_HYDRAULIKSTATIONS_NR )
  THEN
    refMK REF= apgMKHydraulikstation[wpHydraulikstationNr];
  END_IF
END_IF

//-------------------------------------------------------------------------------------------------
// ANFORDERUNGEN UEBERNEHMEN
//-------------------------------------------------------------------------------------------------
(* Hinweis:
   - Die Faecherwagenstationen melden ihre Anforderungen vor diesem Aufruf ueber M_Anfordern
     und ihre Auftraege ueber M_AuftragFreigabe
   - Uebernehmen und fuer den naechsten Zyklus loeschen
*)
blHydraulikStarten             := blAnforderungHydraulik;
blUmlaufventilPause            := blAnforderungUmlaufventilPause;
blAnforderungHydraulik         := FALSE;
blAnforderungUmlaufventilPause := FALSE;
wlAktiveAuftraege              := wlAktiveAuftraegeZyklus;
wlAktiveAuftraegeZyklus        := 0;
wlNeueAuftraegeZyklus          := 0;

//-------------------------------------------------------------------------------------------------
// DEAKTIVIEREN
//-------------------------------------------------------------------------------------------------
IF NOT __ISVALIDREF(refMK) THEN
  out_bHydraulikkreislauf_MotorEin        := FALSE;
  out_bHydraulikkreislauf_UmlaufventilAuf := FALSE;
  bpHydraulikLaeuft                       := FALSE;
  RETURN;
END_IF

IF ( refMK.bDeaktivieren ) THEN
  tonlUmlaufventilEin( IN := FALSE );
  out_bHydraulikkreislauf_MotorEin        := FALSE;
  out_bHydraulikkreislauf_UmlaufventilAuf := FALSE;
  bpHydraulikLaeuft                       := FALSE;
  RETURN;
END_IF

//-------------------------------------------------------------------------------------------------
// PROZESS
//-------------------------------------------------------------------------------------------------
(* Hinweis:
   - Motor laeuft, solange eine Station eine hydraulische Bewegung anfordert
   - Umlaufventil nach wgTimeHydraulikUmlaufEin schalten; eine Station kann es zwischen zwei
     direkt folgenden Bewegungen kurz zuruecknehmen (Pause)
*)
out_bHydraulikkreislauf_MotorEin := blHydraulikStarten;

tonlUmlaufventilEin( IN := out_bHydraulikkreislauf_MotorEin AND NOT blUmlaufventilPause,
                     PT := WORD_TO_TIME( wgTimeHydraulikUmlaufEin * cUMRECHNUNG_MILLISEKUNDEN_SEKUNDEN ) );

out_bHydraulikkreislauf_UmlaufventilAuf := tonlUmlaufventilEin.Q;

//-------------------------------------------------------------------------------------------------
// AUSGAENGE
//-------------------------------------------------------------------------------------------------
bpHydraulikLaeuft :=     out_bHydraulikkreislauf_MotorEin
                     AND out_bHydraulikkreislauf_UmlaufventilAuf
                     AND in_bMotorschuetz_Hydraulikkreislauf_OK;

//-------------------------------------------------------------------------------------------------
// MELDUNGEN
//-------------------------------------------------------------------------------------------------
WatchIo( NOT in_bMotorschuetz_Hydraulikkreislauf_OK, refMK.wMeldungsNummer );
END_FUNCTION_BLOCK
